INTERFACE ITF_Buffer5

METHOD Aborted : BOOL
VAR_INPUT
END_VAR
END_METHOD

METHOD Aborting : BOOL
VAR_INPUT
END_VAR
END_METHOD

METHOD Clearing : BOOL
VAR_INPUT
END_VAR
END_METHOD

METHOD Execute : BOOL
VAR_INPUT
END_VAR
END_METHOD

METHOD Held : BOOL
VAR_INPUT
END_VAR
END_METHOD

METHOD Holding : BOOL
VAR_INPUT
END_VAR
END_METHOD

METHOD Idle : BOOL
VAR_INPUT
END_VAR
END_METHOD

METHOD Resetting : BOOL
VAR_INPUT
END_VAR
END_METHOD

METHOD Starting : BOOL
VAR_INPUT
END_VAR
END_METHOD

METHOD Stopped : BOOL
VAR_INPUT
END_VAR
END_METHOD

METHOD Stopping : BOOL
VAR_INPUT
END_VAR
END_METHOD

METHOD Suspended : BOOL
VAR_INPUT
END_VAR
END_METHOD

METHOD Suspending : BOOL
VAR_INPUT
END_VAR
END_METHOD

METHOD Unholding : BOOL
VAR_INPUT
END_VAR
END_METHOD

METHOD Unsuspending : BOOL
VAR_INPUT
END_VAR
END_METHOD

END_INTERFACE

(* stored: Version 1.1.0.1
   Itf ITF_Buffer5: Id {a881b87c-3a5a-4a95-ba6e-f165b156f503}
   Folder Methods: Id {41da5b41-acf7-4733-91cb-ca533afdc53a}
   Method Aborted: Id {39c6bab9-b1a6-4118-a35b-3771df847f4a}
   Method Aborting: Id {d9e3478d-fcb2-4f74-8219-e6fa7f0f0718}
   Method Clearing: Id {eca19e3f-bf29-43cc-8be1-a4a3920e913d}
   Method Execute: Id {75f539ca-e13b-4ba7-bd6c-0a0f4c8ff602}
   Method Held: Id {0e12e719-fc7e-40d3-ad61-373f103b4dff}
   Method Holding: Id {25c41b9c-9d63-4031-be0a-69de24ca0d19}
   Method Idle: Id {486461dd-8983-4f29-830d-1cc54ec9378f}
   Method Resetting: Id {9d87d0da-c798-49f4-b40c-cc4efa8d1476}
   Method Starting: Id {9d7a17da-3477-4482-bf5e-119626016ec2}
   Method Stopped: Id {dbf1dc7a-0a1f-4525-8633-e90e79cdc2fc}
   Method Stopping: Id {975a4a9d-c181-43e3-852f-369ec13e6fbe}
   Method Suspended: Id {09a088bc-bf19-4450-8486-a538faffb8b3}
   Method Suspending: Id {c13b29a9-b52e-4638-aa3e-91448278b7aa}
   Method Unholding: Id {6c9c7e32-6bf4-46de-97ab-756a85457139}
   Method Unsuspending: Id {49999f61-062c-4f1a-8f73-18ae5ca2be40} *)
